(*
SPDX-FileCopyrightText: © 2026 Oleksandr Tiutyk <trofimich@gmail.com>
SPDX-License-Identifier: MIT
License: https://opensource.org/license/mit
*)

(*!
<summary>Identifies the current queue cleanup test phase.</summary>
*)
{attribute 'qualified_only'}
{attribute 'strict'}
TYPE QUEUE_CLEANUP_TEST_PHASE :
(
	//! <summary>Drive the original failure and child cleanup.</summary>
	FAILURE_RUN,
	//! <summary>Drive the same queue after Reset without a child failure.</summary>
	REUSE_RUN,
	//! <summary>Advance the stopped queue once to check that release is not retried.</summary>
	OBSERVE_FAILED_RELEASE
);
END_TYPE

(* stored: Version 1.1.0.1
   DUT QUEUE_CLEANUP_TEST_PHASE: Id {546ec53b-f1f2-482b-83b6-d303bf463d27} *)
